(* IEC 61131-3 sources: T4Exjobb/Sigma/Stations/MachineControl/MachineControl/Class/_TCPIP_CLIENT (part 2) *)

    (*===============================================================================================*)
    MTERROR_NOFCT: // - CREATE TASK NEEDS A VALID TASK FUNCTION
    (*===============================================================================================*)
      co_SigCLib.StrCpy(pErrTxt, "MTERROR_NOFCT");

    (*===============================================================================================*)
    MTERROR_FCTNOTINMEM: // - CREATE TASK NEEDS A TASK FUNCTION PLACED IN LASAL CODE MEMORY
    (*===============================================================================================*)
      co_SigCLib.StrCpy(pErrTxt, "MTERROR_FCTNOTINMEM");

    (*===============================================================================================*)
    MTERROR_WRONGPRIOR: // - CREATE TASK ONLY SUPPORTS PRIORS FROM 1 .. 14
    (*===============================================================================================*)
      co_SigCLib.StrCpy(pErrTxt, "MTERROR_WRONGPRIOR");

    (*===============================================================================================*)
    MTERROR_STACK: // - CREATE TASK ONLY SUPPORT SATCK SIZE LOWER THAN 0x4000
    (*===============================================================================================*)
      co_SigCLib.StrCpy(pErrTxt, "MTERROR_STACK");

    (*===============================================================================================*)
    MTERROR_NAME: // - CREATE TASK, MAILBOX OR SEMAPHORE NEEDS A VALID NAME
    (*===============================================================================================*)
      co_SigCLib.StrCpy(pErrTxt, "MTERROR_NAME");

    (*===============================================================================================*)
    MTERROR_NAMEUSED: // - CREATE TASK, MAILBOX OR SEMAPHORE NAME ALREADY IN USE
    (*===============================================================================================*)
      co_SigCLib.StrCpy(pErrTxt, "MTERROR_NAMEUSED");

    (*===============================================================================================*)
    MTERROR_HANDLE: // - HANDLE NOT FOUND IN OS-LIST => NOT VALID
    (*===============================================================================================*)
      co_SigCLib.StrCpy(pErrTxt, "MTERROR_HANDLE");

    (*===============================================================================================*)
    MTERROR_NOTALLOWED: // - MT-FUNCTION NOT ALLOWED IN THIS TASK CONTEXT
    (*===============================================================================================*)
      co_SigCLib.StrCpy(pErrTxt, "MTERROR_NOTALLOWED");

    (*===============================================================================================*)
    MTERROR_MESSAGESIZE: // - MAILBOX NEED A VALID MESSAGE SIZE
    (*===============================================================================================*)
      co_SigCLib.StrCpy(pErrTxt, "MTERROR_MESSAGESIZE");

    (*===============================================================================================*)
    MTERROR_DATA: // - POINTER TO DATA IS NOT VALID
    (*===============================================================================================*)
      co_SigCLib.StrCpy(pErrTxt, "MTERROR_DATA");

    (*===============================================================================================*)
    MTERROR_PTR: // - INVALID POINTER, PARAMETER OR INTERNAL
    (*===============================================================================================*)
      co_SigCLib.StrCpy(pErrTxt, "MTERROR_PTR");

    (*===============================================================================================*)
    MTERROR_TASKID: // - INVALID TASK ID, ID NOT FOUND
    (*===============================================================================================*)
      co_SigCLib.StrCpy(pErrTxt, "MTERROR_TASKID");

    (*===============================================================================================*)
    MTERROR_NOTASK: // - TASK DOES NOT EXIST
    (*===============================================================================================*)
      co_SigCLib.StrCpy(pErrTxt, "MTERROR_NOTASK");

    (*===============================================================================================*)
    MTERROR_NOIFFNC: // - INTERFACE FUNCTION IS NOT AVAILABLE
    (*===============================================================================================*)
      co_SigCLib.StrCpy(pErrTxt, "MTERROR_NOIFFNC");

    (*===============================================================================================*)
    else // - UNKNOWN ERROR CODE
    (*===============================================================================================*)
      co_SigCLib.StrCpy(pErrTxt, "MTERROR_UNKNOWN");

  end_case;

END_FUNCTION

FUNCTION _TCPIP_CLIENT::AP_TaskCreate
VAR_INPUT
  pTaskName 	: ^CHAR;
  pCallback 	: ^void;
END_VAR
VAR_OUTPUT
  Retcode 	  : DINT;
END_VAR

  Retcode := TCP_CLT_NO_ERROR;

  AP_TaskHandle := co_MultiTask.CREATETHREAD(pCallback, AP_TaskPriority, 0x4000, MT_TASK_SAVETHIS, this, pTaskName);
  if (AP_TaskHandle = NIL) then
    Retcode := TCP_CLT_ERR_TASK_CREATE;
  end_if;

END_FUNCTION

FUNCTION __CDECL _TCPIP_CLIENT::AP_TaskCallback
VAR_INPUT
#pragma warning (disable: 0073)
  Param0 	: ^void;
#pragma warning (default: 0073)
END_VAR

  while 1 do
    CyclicCall();
    AP_TaskDelay(AP_TaskTime);
  end_while;

END_FUNCTION

FUNCTION _TCPIP_CLIENT::AP_TaskDelay
VAR_INPUT
  udTaskDelay 	: UDINT;
END_VAR

  if (bdStatus.SalamanderOS = true) then
    OSSD_DELAY(pCIL_DEBUG, udTaskDelay);
  else
    co_MultiTask.TASKDELAY(udTaskDelay);
  end_if;

END_FUNCTION

FUNCTION _TCPIP_CLIENT::AP_SemaCreate
VAR_INPUT
  pSemaName 	: ^CHAR;
  Index 	    : DINT;
END_VAR
VAR_OUTPUT
  Retcode 	: DINT;
END_VAR

  Retcode := TCP_CLT_NO_ERROR;

  if (pSemaName <> NIL) then
    case Index of
      (*=================================================================================*)
      0:
      (*=================================================================================*)
        AP_SemaHandle1 := co_MultiTask.CREATESEMAPHORE(MTSEMATYPE_MUTEX, 1, 0, pSemaName);
        if (AP_SemaHandle1 = NIL) then
          Retcode := TCP_CLT_ERR_SEMA_CREATE;
        end_if;

      (*=================================================================================*)
      1:
      (*=================================================================================*)
        AP_SemaSockOpt := co_MultiTask.CREATESEMAPHORE(MTSEMATYPE_MUTEX, 1, 0, pSemaName);
        if (AP_SemaSockOpt = NIL) then
          Retcode := TCP_CLT_ERR_SEMA_CREATE;
        end_if;

      (*=================================================================================*)
      else
      (*=================================================================================*)
        Retcode := TCP_CLT_ERR_SEMA_INVALID_IDX;

    end_case;
  else
    Retcode := TCP_CLT_ERR_SEMA_INVALID_NAME;
  end_if;

END_FUNCTION

FUNCTION _TCPIP_CLIENT::AP_SemaWait
VAR_INPUT
  SemaHandle 	: MT_SEMAHANDLE;
END_VAR

  if (SemaHandle <> NIL) then
    co_MultiTask.WAIT(SemaHandle);
  end_if;

END_FUNCTION

FUNCTION _TCPIP_CLIENT::AP_SemaSignal
VAR_INPUT
  SemaHandle 	: MT_SEMAHANDLE;
END_VAR

  if (SemaHandle <> NIL) then
    co_MultiTask.SIGNAL(SemaHandle);
  end_if;

END_FUNCTION

FUNCTION _TCPIP_CLIENT::DelConnIntern
VAR_INPUT
  pDelConn 	  : ^_CONNECTION;
END_VAR
VAR
	pSearchConn : ^_CONNECTION;
END_VAR

  if (pDelConn <> NIL) then

    AP_SemaWait(AP_SemaHandle1);

    if (pDelConn^.pNextConn = pDelConn) then
      // - ONE ACTIVE CONNECTION
    else
      pSearchConn := pDelConn;
      while pSearchConn^.pNextConn <> pDelConn do
        pSearchConn := pSearchConn^.pNextConn;
      end_while;
      pSearchConn^.pNextConn := pDelConn^.pNextConn;
      pActConn := pDelConn^.pNextConn;
      bdStatus.InhibNextConn := true;
    end_if;

    ConnInfoCallback(pDelConn, TCP_CLT_INFO_DELETED, 0);
    INITConnection(pDelConn);
    AP_SemaSignal(AP_SemaHandle1);

    ActConn -= 1;

  end_if;

END_FUNCTION

FUNCTION VIRTUAL GLOBAL _TCPIP_CLIENT::AddConnectionSSL
VAR_INPUT
  pIPAddress 	                  : ^CHAR;
  pCACertPEMFilename 	          : ^CHAR;
  pClientCertChainPEMFilename 	: ^CHAR;
  pClientCertKeyPEMFilename 	  : ^CHAR;
  pKeyDecryptPwd 	              : ^CHAR;
  pCallbackThis 	              : ^void;
  pCallbackMeth 	              : ^void;
  udTimeout 	                  : UDINT;
END_VAR
VAR_OUTPUT
  dHandle 	                    : DINT;
END_VAR
VAR
	dRet                          : DINT;
END_VAR

  dHandle := 0;

  if (usInit > 0) then
    if (bdStatus.CIL_ssl_user = true) then
      if (bdStatus.ErrMem = false) then
        dRet := CheckParaConnSSL(pCACertPEMFilename, pClientCertChainPEMFilename, pClientCertKeyPEMFilename, pKeyDecryptPwd);
        if (dRet = TCP_CLT_NO_ERROR) then
          dRet := CheckParaConnTCP(pIPAddress, pCallbackThis, pCallbackMeth);
          if (dRet = TCP_CLT_NO_ERROR) then

            dHandle := AddConnIntern(pIPAddress,
                                     pCACertPEMFilename,
                                     pClientCertChainPEMFilename,
                                     pClientCertKeyPEMFilename,
                                     pKeyDecryptPwd,
                                     pCallbackThis,
                                     pCallbackMeth,
                                     udTimeout,
                                     true);

          else
            LastError := dRet;
          end_if;
        else
          LastError := dRet;
        end_if;
      else
        LastError := TCP_CLT_ERR_CONN_MEMORY;
      end_if;
    else
      LastError := TCP_CLT_ERR_NO_SSL_INTERFACE;
    end_if;
  else
    LastError := TCP_CLT_ERR_MAIN_INIT;
  end_if;

END_FUNCTION

FUNCTION _TCPIP_CLIENT::AddConnIntern
VAR_INPUT
  pIPAddress 	                  : ^CHAR;
  pCACertPEMFilename 	          : ^CHAR;
  pClientCertChainPEMFilename 	: ^CHAR;
  pClientCertKeyPEMFilename 	  : ^CHAR;
  pKeyDecryptPwd 	              : ^CHAR;
  pCallbackThis 	              : ^void;
  pCallbackMeth 	              : ^void;
  udTimeout 	                  : UDINT;
  ConnSSL 	                    : BOOL;
END_VAR
VAR_OUTPUT
  dHandle 	                    : DINT;
END_VAR
VAR
  pFirstConn                    : ^_CONNECTION;
  pNewConn                      : ^_CONNECTION;
  pSearchConn                   : ^_CONNECTION;
  i                             : USINT;
END_VAR

  dHandle := 0;

  if (pIPAddress = NIL) | (pConnectionBuffer = NIL) | (Control = _STATE_ERROR_CREATING_MUTEX) | (Control = _STATE_ERROR_ALLOCATING_MEMORY) then
    return;
  end_if;

  if (ActConn < MaxConn) then

    AP_SemaWait(AP_SemaHandle1);

    for i := 0 to (MaxConn-1) do
      pFirstConn := pConnectionBuffer + (i * sizeof(_CONNECTION));
      if (pFirstConn^.bInUse = true) then
        exit;
      else
        pFirstConn := NIL;
      end_if;
    end_for;

    for i := 0 to (MaxConn-1) do
      pNewConn := pConnectionBuffer + (i * sizeof(_CONNECTION));
      if (pNewConn^.bInUse = false) then
        exit;
      end_if;
    end_for;

    pNewConn^.bInUse          := true;
    pNewConn^.udTimeout       := udTimeout;
    pNewConn^.pCallbackThis   := pCallbackThis;
    pNewConn^.pCallbackMeth   := pCallbackMeth;
    pNewConn^.FSM_TCP         := _STATE_IDLE;
    pNewConn^.ConnSockOpt     := MainSockOpt;
    pNewConn^.KeepAlivePara   := KeepAlivePara;
    pNewConn^.CloseSocketType := CloseSocketType;
    co_SigCLib.StrCpy(#pNewConn^.szIPAddress[0], pIPAddress);
    pNewConn^.bdSettings.SockOptChanged := true;

    if (ConnSSL = true) then
      pNewConn^.bdSettings.ConnSSL := true;
      if (pCACertPEMFilename <> NIL) then
        co_SigCLib.StrCpy(#pNewConn^.szCACertPEMFileName[0], pCACertPEMFilename);
      end_if;
      if (pClientCertChainPEMFilename <> NIL) then
        co_SigCLib.StrCpy(#pNewConn^.szClientCertChainPEMFilename[0], pClientCertChainPEMFilename);
      end_if;
      if (pClientCertKeyPEMFilename <> NIL) then
        co_SigCLib.StrCpy(#pNewConn^.szClientCertKeyPEMFilename[0], pClientCertKeyPEMFilename);
      end_if;
      if (pKeyDecryptPwd <> NIL) then
        co_SigCLib.StrCpy(#pNewConn^.szKeyDecryptPwd[0], pKeyDecryptPwd);
      end_if;
    end_if;

    if (pFirstConn = NIL) then
      pNewConn^.pNextConn := pNewConn;
    else
      pSearchConn := pFirstConn;
      while (pSearchConn^.pNextConn <> pFirstConn) do
        pSearchConn := pSearchConn^.pNextConn;
      end_while;
      pNewConn^.pNextConn    := pFirstConn;
      pSearchConn^.pNextConn := pNewConn;
    end_if;

    dHandle := pNewConn$DINT;
    ActConn += 1;

    AP_SemaSignal(AP_SemaHandle1);

  else
    LastError := TCP_CLT_ERR_MAX_CONN;
  end_if;

END_FUNCTION

FUNCTION _TCPIP_CLIENT::CheckParaConnSSL
VAR_INPUT
  pCACertPEMFilename 	          : ^CHAR;
  pClientCertChainPEMFilename 	: ^CHAR;
  pClientCertKeyPEMFilename 	  : ^CHAR;
  pKeyDecryptPwd 	              : ^CHAR;
END_VAR
VAR_OUTPUT
  Retcode 	                    : DINT;
END_VAR

  Retcode := TCP_CLT_NO_ERROR;

  if (pClientCertChainPEMFilename <> NIL) then
    if (pClientCertKeyPEMFilename = NIL) then
      Retcode := TCP_CLT_ERR_INVALID_PARA_SSL;
    end_if;
  end_if;

  if (pClientCertKeyPEMFilename <> NIL) then
    if (pClientCertChainPEMFilename = NIL) then
      Retcode := TCP_CLT_ERR_INVALID_PARA_SSL;
    end_if;
  end_if;

  if (pKeyDecryptPwd <> NIL) then
    if (pClientCertChainPEMFilename = NIL) then
      Retcode := TCP_CLT_ERR_INVALID_PARA_SSL;
    end_if;
    if (pClientCertKeyPEMFilename = NIL) then
      Retcode := TCP_CLT_ERR_INVALID_PARA_SSL;
    end_if;
  end_if;

END_FUNCTION

FUNCTION _TCPIP_CLIENT::FindFirstConn
VAR_OUTPUT
  pFirstConn 	: ^_CONNECTION;
END_VAR
VAR
	i           : USINT;
  pSearchConn : ^_CONNECTION;
END_VAR

  pFirstConn := NIL;

  for i := 0 to (MaxConn-1) do
    pSearchConn := pConnectionBuffer + (i * sizeof(_CONNECTION));
    if (pSearchConn^.bInUse = true) then
      pFirstConn := pSearchConn;
    end_if;
  end_for;

END_FUNCTION

FUNCTION _TCPIP_CLIENT::CheckParaConnTCP
VAR_INPUT
  pIPAddress 	    : ^CHAR;
  pCallbackThis 	: ^void;
  pCallbackMeth 	: ^void;
END_VAR
VAR_OUTPUT
  Retcode 	      : DINT;
END_VAR
VAR
	udStrLen        : UDINT;
END_VAR

  Retcode := TCP_CLT_NO_ERROR;

  if (pIPAddress = NIL) then
    Retcode := TCP_CLT_ERR_INVALID_PARA_TCP;
  else
    udStrLen := co_SigCLib.StrLen(pIPAddress);
    if (udStrLen = 0) then
      Retcode := TCP_CLT_ERR_INVALID_PARA_TCP;
    end_if;
  end_if;

//  if (pCallbackThis = NIL) then
//    Retcode := TCP_CLT_ERR_INVALID_PARA_TCP;
//  end_if;
//
//  if (pCallbackMeth = NIL) then
//    Retcode := TCP_CLT_ERR_INVALID_PARA_TCP;
//  end_if;

END_FUNCTION

FUNCTION GLOBAL _TCPIP_CLIENT::GetLastError
VAR_OUTPUT
  Retcode 	: DINT;
END_VAR

  Retcode := LastError;

END_FUNCTION

FUNCTION GLOBAL _TCPIP_CLIENT::InstallConnErrCallback
VAR_INPUT
  dHandle 	      : DINT;
  pCallbackThis 	: ^void;
  pCallbackMeth 	: ^void;
END_VAR
VAR_OUTPUT
  Retcode 	      : DINT;
END_VAR
VAR
	pConn           : ^_CONNECTION;
END_VAR

  Retcode := TCP_CLT_NO_ERROR;

  if (CheckHandleValid(dHandle) = true) then
    if (pCallbackThis <> NIL) & (pCallbackMeth <> NIL) then
      pConn := dHandle$^_CONNECTION;
      pConn^.pErrCallbackThis := pCallbackThis;
      pConn^.pErrCallbackMeth := pCallbackMeth;
    else
      Retcode := TCP_CLT_ERR_INVALID_POINTER;
    end_if;
  else
    Retcode := TCP_CLT_INVALID_HANDLE;
  end_if;

END_FUNCTION

FUNCTION _TCPIP_CLIENT::ErrCallback
VAR_INPUT
#pragma warning (disable: 0073)
  FSM_TCP 	: _FSM_TCP_USER;
  ErrGroup 	: DINT;
  ErrCode 	: DINT;
#pragma warning (default: 0073)
END_VAR

END_FUNCTION

FUNCTION _TCPIP_CLIENT::ConnErrCallback
VAR_INPUT
  pConn 	  : ^_CONNECTION;
  ErrGroup 	: DINT;
  ErrCode 	: DINT;
END_VAR
VAR_OUTPUT
  Retcode 	: DINT;
END_VAR
VAR
	pTmpThis  : ^void;
END_VAR

  Retcode := TCP_CLT_NO_ERROR;

  if (pConn <> NIL) then
    if (pConn^.pErrCallbackThis <> NIL) & (pConn^.pErrCallbackMeth <> NIL) then
      pTmpThis := this;
      this$^void := pConn^.pErrCallbackThis;
      #pragma warning(disable: 137);
      pConn^.pErrCallbackMeth$ErrCallback(pConn^.FSM_TCP, ErrGroup, ErrCode);
      #pragma warning(default: 137);
      this$^void := pTmpThis;
    end_if;
  else
    Retcode := TCP_CLT_INVALID_HANDLE;
  end_if;

END_FUNCTION

FUNCTION VIRTUAL GLOBAL _TCPIP_CLIENT::ReadMainParameter
VAR_INPUT
  Cmd 	      : DINT;
  SubCmd 	    : DINT;
  pParaValue 	: ^DINT;
END_VAR
VAR_OUTPUT
  Retcode 	  : DINT;
END_VAR

  Retcode := TCP_CLT_NO_ERROR;

  if (usInit > 0) then
    case Cmd of
      (*================================================================*)
      TCPCLT_CMD_SETSOCKOPT:
      (*================================================================*)
        case SubCmd of
          (*==================================================*)
          TCPCLT_SOCKOPT_NAGLE:
          (*==================================================*)
            if (MainSockOpt.Nagle = false) then
              pParaValue^ := 0;
            else
              pParaValue^ := 1;
            end_if;
          (*==================================================*)
          TCPCLT_SOCKOPT_KEEPALIVE:
          (*==================================================*)
            if (MainSockOpt.KeepAlive = false) then
              pParaValue^ := 0;
            else
              pParaValue^ := 1;
            end_if;
          (*==================================================*)
          TCPCLT_SOCKOPT_DELAYEDACK:
          (*==================================================*)
            if (MainSockOpt.DelayedAck = false) then
              pParaValue^ := 0;
            else
              pParaValue^ := 1;
            end_if;
          (*==================================================*)
          else // - INVALID SUB COMMAND
          (*==================================================*)
            Retcode := TCP_CLT_ERR_SET_PARA_INVALID_SUB_CMD;
        end_case;

      (*================================================================*)
      TCPCLT_CMD_TASKPRIO:
      (*================================================================*)
        case SubCmd of
          (*==================================================*)
          TCPCLT_SUB_CMD_TASKPRIO:
          (*==================================================*)
            pParaValue^ := AP_TaskPriority$DINT;
          (*==================================================*)
          else // - INVALID SUB COMMAND
          (*==================================================*)
            Retcode := TCP_CLT_ERR_SET_PARA_INVALID_SUB_CMD;
        end_case;

      (*================================================================*)
      TCPCLT_CMD_KEEPALIVEPARA:
      (*================================================================*)
        case SubCmd of
          (*==================================================*)
          TCPCLT_KEEPALIVE_KEEPIDLE:
          (*==================================================*)
            pParaValue^ := KeepAlivePara.keepIDLE;
          (*==================================================*)
          TCPCLT_KEEPALIVE_KEEPINTVL:
          (*==================================================*)
            pParaValue^ := KeepAlivePara.keepINTVL;
          (*==================================================*)
          TCPCLT_KEEPALIVE_KEEPCNT:
          (*==================================================*)
            pParaValue^ := KeepAlivePara.keepCNT;
          (*==================================================*)
          else // - INVALID SUB COMMAND
          (*==================================================*)
            Retcode := TCP_CLT_ERR_SET_PARA_INVALID_SUB_CMD;
        end_case;

      (*================================================================*)
      TCPCLT_CMD_CLOSESOCKETTYPE:
      (*================================================================*)
        case SubCmd of
          (*==================================================*)
          TCPCLT_CLOSESOCKETTYPE:
          (*==================================================*)
            pParaValue^$UDINT := CloseSocketType;
          (*==================================================*)
          else // - INVALID SUB COMMAND
          (*==================================================*)
            Retcode := TCP_CLT_ERR_SET_PARA_INVALID_SUB_CMD;
        end_case;

      (*================================================================*)
      else // - INVALID COMMAND
      (*================================================================*)
        Retcode := TCP_CLT_ERR_SET_PARA_INVALID_CMD;

    end_case;
  else
    Retcode := TCP_CLT_ERR_MAIN_INIT;
  end_if;

END_FUNCTION

FUNCTION VIRTUAL GLOBAL _TCPIP_CLIENT::ReadConnParameter
VAR_INPUT
  dHandle 	  : DINT;
  Cmd 	      : DINT;
  SubCmd 	    : DINT;
  pParaValue 	: ^DINT;
END_VAR
VAR_OUTPUT
  Retcode 	  : DINT;
END_VAR
VAR
	pConn       : ^_CONNECTION;
END_VAR

  Retcode := TCP_CLT_NO_ERROR;

  if (CheckHandleValid(dHandle) = true) then
    pConn := dHandle$^_CONNECTION;
    case Cmd of
      (*================================================================*)
      TCPCLT_CMD_SETSOCKOPT:
      (*================================================================*)
        if (pConn^.bdSettings.ConnSSL = true) then
          Retcode := TCP_CLT_ERR_SET_PARA_CMD_NOT_SUPPORTED;
        else
          case SubCmd of
            (*==================================================*)
            TCPCLT_SOCKOPT_NAGLE:
            (*==================================================*)
              if (pConn^.ConnSockOpt.Nagle = false) then
                pParaValue^ := 0;
              else
                pParaValue^ := 1;
              end_if;
            (*==================================================*)
            TCPCLT_SOCKOPT_KEEPALIVE:
            (*==================================================*)
              if (pConn^.ConnSockOpt.KeepAlive = false) then
                pParaValue^ := 0;
              else
                pParaValue^ := 1;
              end_if;
            (*==================================================*)
            TCPCLT_SOCKOPT_DELAYEDACK:
            (*==================================================*)
              if (pConn^.ConnSockOpt.DelayedAck = false) then
                pParaValue^ := 0;
              else
                pParaValue^ := 1;
              end_if;
            (*==================================================*)
            else // - INVALID SUB COMMAND
            (*==================================================*)
              Retcode := TCP_CLT_ERR_SET_PARA_INVALID_SUB_CMD;
          end_case;
        end_if;

      (*================================================================*)
      TCPCLT_CMD_KEEPALIVEPARA:
      (*================================================================*)
        if (pConn^.bdSettings.ConnSSL = true) then
          Retcode := TCP_CLT_ERR_SET_PARA_CMD_NOT_SUPPORTED;
        else
          case SubCmd of
            (*==================================================*)
            TCPCLT_KEEPALIVE_KEEPIDLE:
            (*==================================================*)
              pParaValue^ := pConn^.KeepAlivePara.keepIDLE;
            (*==================================================*)
            TCPCLT_KEEPALIVE_KEEPINTVL:
            (*==================================================*)
              pParaValue^ := pConn^.KeepAlivePara.keepINTVL;
            (*==================================================*)
            TCPCLT_KEEPALIVE_KEEPCNT:
            (*==================================================*)
              pParaValue^ := pConn^.KeepAlivePara.keepCNT;
            (*==================================================*)
            else // - INVALID SUB COMMAND
            (*==================================================*)
              Retcode := TCP_CLT_ERR_SET_PARA_INVALID_SUB_CMD;
          end_case;
        end_if;

      (*================================================================*)
      TCPCLT_CMD_CLOSESOCKETTYPE:
      (*================================================================*)
        if (pConn^.bdSettings.ConnSSL = true) then
          Retcode := TCP_CLT_ERR_SET_PARA_CMD_NOT_SUPPORTED;
        else
          case SubCmd of
            (*==================================================*)
            TCPCLT_CLOSESOCKETTYPE:
            (*==================================================*)
              pParaValue^$UDINT := pConn^.CloseSocketType;
            (*==================================================*)
            else // - INVALID SUB COMMAND
            (*==================================================*)
              Retcode := TCP_CLT_ERR_SET_PARA_INVALID_SUB_CMD;
          end_case;
        end_if;

      (*================================================================*)
      else // - INVALID COMMAND
      (*================================================================*)
        Retcode := TCP_CLT_ERR_SET_PARA_INVALID_CMD;

    end_case;
  else
    Retcode := TCP_CLT_INVALID_HANDLE;
  end_if;

END_FUNCTION

FUNCTION GLOBAL _TCPIP_CLIENT::InstallConnInfoCallback
VAR_INPUT
  dHandle 	      : DINT;
  pCallbackThis 	: ^void;
  pCallbackMeth 	: ^void;
END_VAR
VAR_OUTPUT
  Retcode 	      : DINT;
END_VAR
VAR
	pConn           : ^_CONNECTION;
END_VAR

  Retcode := TCP_CLT_NO_ERROR;

  if (CheckHandleValid(dHandle) = true) then
    if (pCallbackThis <> NIL) & (pCallbackMeth <> NIL) then
      pConn := dHandle$^_CONNECTION;
      pConn^.pInfoCallbackThis := pCallbackThis;
      pConn^.pInfoCallbackMeth := pCallbackMeth;
    else
      Retcode := TCP_CLT_ERR_INVALID_POINTER;
    end_if;
  else
    Retcode := TCP_CLT_INVALID_HANDLE;
  end_if;

END_FUNCTION

FUNCTION _TCPIP_CLIENT::InfoCallback
VAR_INPUT
#pragma warning (disable: 0073)
  FSM_TCP 	: _FSM_TCP_USER;
  InfoPara1 	: DINT;
  InfoPara2 	: DINT;
#pragma warning (default: 0073)
END_VAR

END_FUNCTION

FUNCTION _TCPIP_CLIENT::ConnInfoCallback
VAR_INPUT
  pConn 	    : ^_CONNECTION;
  InfoPara1 	: DINT;
  InfoPara2 	: DINT;
END_VAR
VAR_OUTPUT
  Retcode 	  : DINT;
END_VAR
VAR
	pTmpThis    : ^void;
END_VAR

  Retcode := TCP_CLT_NO_ERROR;

  if (pConn <> NIL) then
    if (pConn^.pInfoCallbackThis <> NIL) & (pConn^.pInfoCallbackMeth <> NIL) then
      pTmpThis := this;
      this$^void := pConn^.pInfoCallbackThis;
      #pragma warning(disable: 137);
      pConn^.pInfoCallbackMeth$InfoCallback(pConn^.FSM_TCP, InfoPara1, InfoPara2);
      #pragma warning(default: 137);
      this$^void := pTmpThis;
    end_if;
  else
    Retcode := TCP_CLT_INVALID_HANDLE;
  end_if;

END_FUNCTION

FUNCTION _TCPIP_CLIENT::Callback
VAR_INPUT
#pragma warning (disable: 0073)
  pData   : ^void;
  udSize  : UDINT;
#pragma warning (default: 0073)
END_VAR

END_FUNCTION

FUNCTION _TCPIP_CLIENT::AP_NReadAvailable
VAR_INPUT
  pConn 	: ^_CONNECTION;
END_VAR
VAR_OUTPUT
  Retcode 	: DINT;
END_VAR

  if (pConn <> NIL) then
    if (pConn^.bdSettings.ConnSSL = false) then
      Retcode := OS_TCP_USER_NREAD_AVAILABLE(pConn^.dSocket);
    else
      Retcode := cSizeOfTXBuffer$DINT;
    end_if;
  else
    Retcode := TCP_CLT_INVALID_HANDLE;
  end_if;

END_FUNCTION

FUNCTION VIRTUAL GLOBAL _TCPIP_CLIENT::GetSetting
VAR_INPUT
  Index 	: DINT;
  pSetting 	: ^DINT;
END_VAR
VAR_OUTPUT
  Retcode 	: DINT;
END_VAR

  Retcode := 0;

  case Index of

    (*============================================================================*)
    TCPCLT_GET_SETTING_PORT:
    (*============================================================================*)
      pSetting^ := cPort;

    (*============================================================================*)
    TCPCLT_GET_SETTING_BUFSIZE:
    (*============================================================================*)
      pSetting^ := cSizeOfTXBuffer$DINT;

    (*============================================================================*)
    TCPCLT_GET_SETTING_MAXCONN:
    (*============================================================================*)
      pSetting^ := cMaxConnections;

    (*============================================================================*)
    TCPCLT_GET_SETTING_CONFIG:
    (*============================================================================*)
      pSetting^ := cConfig;

    (*============================================================================*)
    else
    (*============================================================================*)
      Retcode := -1;

  end_case;

END_FUNCTION
